FUNCTION_BLOCK FB_VirtualCylinder
VAR_OUTPUT
    Position : DINT; // 0 = home, 100 = forward limit
END_VAR

METHOD FollowStroke
VAR_INPUT
    Forward : BOOL;
END_VAR
IF Forward THEN
    Position := MIN(100, Position + 1);
ELSE
    Position := MAX(0, Position - 1);
END_IF
END_METHOD

METHOD Home
Position := 0;
END_METHOD

END_FUNCTION_BLOCK

(* stored: Version 1.1.0.1, ProductVersion 3.1.4024.53
   POU FB_VirtualCylinder: Id {52592E20-A431-4FDA-93CC-000000000007}
   Method FollowStroke: Id {52592E20-A431-4FDA-93CC-000000000005}
   Method Home: Id {52592E20-A431-4FDA-93CC-000000000006} *)
